(* IEC 61131-3 sources: plcassist-cli/packages/volt-lsp-iec/test-corpus/CodesysTestProject/Device/Plc Logic/Application/Library Manager/(unresolved)/cmperrors2 interfaces, 1 file *)

(* ---- ERRORS.gvl ---- *)
VAR_GLOBAL
	ERR_OK : UDINT := 16#0;
	ERR_FAILED : UDINT := 16#1;
	ERR_PARAMETER : UDINT := 16#2;
	ERR_NOTINITIALIZED : UDINT := 16#3;
	ERR_VERSION : UDINT := 16#4;
	ERR_TIMEOUT : UDINT := 16#5;
	ERR_NOBUFFER : UDINT := 16#6;
	ERR_PENDING : UDINT := 16#A;
	ERR_NUMPENDING : UDINT := 16#B;
	ERR_NOTIMPLEMENTED : UDINT := 16#C;
	ERR_INVALIDID : UDINT := 16#D;
	ERR_OVERFLOW : UDINT := 16#E;
	ERR_BUFFERSIZE : UDINT := 16#F;
	ERR_NO_OBJECT : UDINT := 16#10;
	ERR_NOMEMORY : UDINT := 16#11;
	ERR_DUPLICATE : UDINT := 16#12;
	ERR_MEMORY_OVERWRITE : UDINT := 16#13;
	ERR_INVALID_HANDLE : UDINT := 16#14;
	ERR_END_OF_OBJECT : UDINT := 16#15;
	ERR_NO_CHANGE : UDINT := 16#16;
	ERR_INVALID_INTERFACE : UDINT := 16#17;
	ERR_NOT_SUPPORTED : UDINT := 16#18;
	ERR_NO_ACCESS_RIGHTS : UDINT := 16#19;
	ERR_OUT_OF_LIMITS : UDINT := 16#1A;
	ERR_ENTRIES_REMAINING : UDINT := 16#1B;
	ERR_INVALID_SESSION_ID : UDINT := 16#1C;
	ERR_EXCEPTION : UDINT := 16#1D;
	ERR_SIGNATURE_MISMATCH : UDINT := 16#1E;
	ERR_VERSION_MISMATCH : UDINT := 16#1F;
	ERR_TYPE_MISMATCH : UDINT := 16#20;
	ERR_ID_MISMATCH : UDINT := 16#21;
	ERR_NO_CONSISTENCY : UDINT := 16#22;
	ERR_NO_COMM_CYCLE : UDINT := 16#23;
	ERR_DONT_SUSPEND_TASK : UDINT := 16#24;
	ERR_MEMORY_LOCK_FAILED : UDINT := 16#25;
	ERR_LICENSE_MISSING : UDINT := 16#26;
	ERR_OPERATION_DENIED : UDINT := 16#27;
	ERR_DEVICE : UDINT := 16#28;
	ERR_DISK_FULL : UDINT := 16#29;
	ERR_CRC_FAILED : UDINT := 16#30;
	ERR_MEDIA_ERASE : UDINT := 16#31;
	ERR_FILE_ERROR : UDINT := 16#32;
	ERR_NO_RETAIN_MEMORY : UDINT := 16#33;
	ERR_OUT_OF_LIMITS_MIN : UDINT := 16#34;
	ERR_OUT_OF_LIMITS_MAX : UDINT := 16#35;
	ERR_SIZE_MISMATCH : UDINT := 16#36;
	ERR_CALL_AGAIN : UDINT := 16#37;
	ERR_NOTHING_TO_DO : UDINT := 16#38;
	ERR_SECURITY_CHECKS_FAILED : UDINT := 16#39;
	ERR_INVALID_SEQUENCE : UDINT := 16#3A;
	ERR_INVALID_REFERENCE : UDINT := 16#3B;
	ERR_CONVERSION_INCOMPLETE : UDINT := 16#3C;
	ERR_TOO_MANY_RETRIES : UDINT := 16#3D;
	ERR_ALIGNMENT : UDINT := 16#3E;
	ERR_CHANGE_PASSWORD : UDINT := 16#3F;
	ERR_REAUTHENTICATE : UDINT := 16#40;
	ERR_RELOGIN : UDINT := 16#41;
	ERR_INVALID_URL : UDINT := 16#42;
	ERR_INVALID_STATE : UDINT := 16#43;
	ERR_USER_MISMATCH : UDINT := 16#44;
	ERR_NOT_READY_YET : UDINT := 16#45;
	ERR_ACTIVATE_USERMGMT : UDINT := 16#46;
	ERR_NO_USERMGMT : UDINT := 16#47;
	ERR_INVALID_ENCODING : UDINT := 16#48;
	ERR_TARGET_MISMATCH : UDINT := 16#49;
	ERR_CLIENT_IN_RO_MODE : UDINT := 16#4A;
	ERR_LICENSE_EXCEEDED : UDINT := 16#4B;
	ERR_ASYNC_EXCEPTION : UDINT := 16#4C;
	ERR_NO_SIGNATURE : UDINT := 16#4D;
	ERR_PASSWORD_POLICY : UDINT := 16#4E;
	ERR_LICENSE_EXPIRED : UDINT := 16#4F;
	ERR_LICENSE_OCCUPIED : UDINT := 16#50;
	ERR_LICENSE_MAINTENANCE_PERIOD_OUTSIDE : UDINT := 16#51;
	ERR_SOCK_NOTINITIALIZED : UDINT := 16#201;
	ERR_SOCK_NOTSOCKET : UDINT := 16#202;
	ERR_SOCK_AFUNSUPPORTED : UDINT := 16#203;
	ERR_SOCK_PROTOUNSUPPORTED : UDINT := 16#204;
	ERR_SOCK_NOBUFFER : UDINT := 16#205;
	ERR_SOCK_WOULDBLOCK : UDINT := 16#206;
	ERR_SOCK_ADDRINUSE : UDINT := 16#207;
	ERR_SOCK_ADDRNOTAVAILABLE : UDINT := 16#208;
	ERR_SOCK_CONNREFUSED : UDINT := 16#209;
	ERR_SOCK_TIMEDOUT : UDINT := 16#20A;
	ERR_SOCK_HOSTNOTFOUND : UDINT := 16#20B;
	ERR_SOCK_HOSTUNREACHABLE : UDINT := 16#20C;
	ERR_SOCK_ISCONNECTED : UDINT := 16#20D;
	ERR_SOCK_NOTCONNECTED : UDINT := 16#20E;
	ERR_SOCK_SHUTDOWN : UDINT := 16#20F;
	ERR_SOCK_MSGSIZE : UDINT := 16#210;
	ERR_SOCK_CLOSED : UDINT := 16#211;
	ERR_L7_TAG_MISSING : UDINT := 16#300;
	ERR_L7_UNKNOWNCMDGROUP : UDINT := 16#301;
	ERR_L7_UNKNOWNCMD : UDINT := 16#302;
	ERR_L7_INCOMPLETE : UDINT := 16#303;
	ERR_CERT_OK : UDINT := ERR_OK;
	ERR_CERT_UNABLE_TO_GET_ISSUER_CERT : UDINT := 16#701;
	ERR_CERT_UNABLE_TO_GET_CRL : UDINT := 16#702;
	ERR_CERT_UNABLE_TO_DECRYPT_CERT_SIGNATURE : UDINT := 16#703;
	ERR_CERT_UNABLE_TO_DECRYPT_CRL_SIGNATURE : UDINT := 16#704;
	ERR_CERT_UNABLE_TO_DECODE_ISSUER_PUBLIC_KEY : UDINT := 16#705;
	ERR_CERT_SIGNATURE_FAILURE : UDINT := 16#706;
	ERR_CERT_CRL_SIGNATURE_FAILURE : UDINT := 16#707;
	ERR_CERT_NOT_YET_VALID : UDINT := 16#708;
	ERR_CERT_HAS_EXPIRED : UDINT := 16#709;
	ERR_CERT_CRL_NOT_YET_VALID : UDINT := 16#70A;
	ERR_CERT_CRL_HAS_EXPIRED : UDINT := 16#70B;
	ERR_CERT_ERROR_IN_CERT_NOT_BEFORE_FIELD : UDINT := 16#70C;
	ERR_CERT_ERROR_IN_CERT_NOT_AFTER_FIELD : UDINT := 16#70D;
	ERR_CERT_ERROR_IN_CRL_LAST_UPDATE_FIELD : UDINT := 16#70E;
	ERR_CERT_ERROR_IN_CRL_NEXT_UPDATE_FIELD : UDINT := 16#70F;
	ERR_CERT_OUT_OF_MEM : UDINT := 16#710;
	ERR_CERT_DEPTH_ZERO_SELF_SIGNED_CERT : UDINT := 16#711;
	ERR_CERT_SELF_SIGNED_CERT_IN_CHAIN : UDINT := 16#712;
	ERR_CERT_UNABLE_TO_GET_ISSUER_CERT_LOCALLY : UDINT := 16#713;
	ERR_CERT_UNABLE_TO_VERIFY_LEAF_SIGNATURE : UDINT := 16#714;
	ERR_CERT_CHAIN_TOO_LONG : UDINT := 16#715;
	ERR_CERT_REVOKED : UDINT := 16#716;
	ERR_CERT_INVALID_CA : UDINT := 16#717;
	ERR_CERT_PATH_LENGTH_EXCEEDED : UDINT := 16#718;
	ERR_CERT_INVALID_PURPOSE : UDINT := 16#719;
	ERR_CERT_UNTRUSTED : UDINT := 16#71A;
	ERR_CERT_REJECTED : UDINT := 16#71B;
	ERR_CERT_SUBJECT_ISSUER_MISMATCH : UDINT := 16#71C;
	ERR_CERT_AKID_SKID_MISMATCH : UDINT := 16#71D;
	ERR_CERT_AKID_ISSUER_SERIAL_MISMATCH : UDINT := 16#71E;
	ERR_CERT_KEYUSAGE_NO_CERTSIGN : UDINT := 16#71F;
	ERR_CERT_UNABLE_TO_GET_CRL_ISSUER : UDINT := 16#720;
	ERR_CERT_UNHANDLED_CRITICAL_EXTENSION : UDINT := 16#721;
	ERR_CERT_KEYUSAGE_NO_CRL_SIGN : UDINT := 16#722;
	ERR_CERT_UNHANDLED_CRITICAL_CRL_EXTENSION : UDINT := 16#723;
	ERR_CERT_INVALID_NON_CA : UDINT := 16#724;
	ERR_CERT_PROXY_PATH_LENGTH_EXCEEDED : UDINT := 16#725;
	ERR_CERT_KEYUSAGE_NO_DIGITAL_SIGNATURE : UDINT := 16#726;
	ERR_CERT_PROXY_CERTIFICATES_NOT_ALLOWED : UDINT := 16#727;
	ERR_CERT_INVALID_EXTENSION : UDINT := 16#728;
	ERR_CERT_INVALID_POLICY_EXTENSION : UDINT := 16#729;
	ERR_CERT_NO_EXPLICIT_POLICY : UDINT := 16#72A;
	ERR_CERT_DIFFERENT_CRL_SCOPE : UDINT := 16#72B;
	ERR_CERT_UNSUPPORTED_EXTENSION_FEATURE : UDINT := 16#72C;
	ERR_CERT_UNNESTED_RESOURCE : UDINT := 16#72D;
	ERR_CERT_PERMITTED_VIOLATION : UDINT := 16#72E;
	ERR_CERT_EXCLUDED_VIOLATION : UDINT := 16#72F;
	ERR_CERT_SUBTREE_MINMAX : UDINT := 16#730;
	ERR_CERT_UNSUPPORTED_CONSTRAINT_TYPE : UDINT := 16#731;
	ERR_CERT_UNSUPPORTED_CONSTRAINT_SYNTAX : UDINT := 16#732;
	ERR_CERT_UNSUPPORTED_NAME_SYNTAX : UDINT := 16#733;
	ERR_CERT_CRL_PATH_VALIDATION_ERROR : UDINT := 16#734;
	ERR_CERT_APPLICATION_VERIFICATION : UDINT := 16#735;
	ERR_CERT_MISSING : UDINT := 16#736;
	ERR_CERT_UNKNOWN_ERROR : UDINT := 16#737;
	ERR_CERT_UNABLE_TO_GET_ISSUER_CRL : UDINT := 16#738;
	ERR_REDU_TOO_TAGS : UDINT := 16#B00;
	ERR_REDU_MEMORY : UDINT := 16#B01;
	ERR_REDU_CLIENT_CREATION_ERR : UDINT := 16#B02;
END_VAR
